(* IEC 61131-3 sources: PLC-Static-Analysis/modules/plc-rules/src/test/resources/PLCA-Q009/named, 1 file *)

(* ---- switch.st ---- *)
PROGRAM P
VAR
    bDone : BOOL;
END_VAR
VAR CONSTANT
    cSimulation : BOOL := FALSE;
END_VAR
IF cSimulation THEN // PLCA-Q009
    bDone := TRUE;
END_IF
END_PROGRAM
